SUBAPPLICATION Checkbox_TO_AD2_2 (* 2 VT-Checkboxes zu einer Bitmaske zusammenfassen und als AD2 (bidirektional) an einen Consumer weiterreichen (z.B. AOption_AD_DEMUX_2.K). Checkbox 1 -> Bit0, Checkbox 2 -> Bit1. Das vom Consumer zurueckgemeldete Echo (die tatsaechlich aktive Bitmaske) wird wieder auf die beiden Checkboxen zurueckgeschrieben. *)
  (* Standard: 61499-2; Description: Copyright (c) 2026 Meisterschulen am Ostbahnhof This program and the accompanying materials are made available under the terms of the Eclipse Public License 2.0 which is available at https://www.eclipse.org/legal/epl-2.0/ SPDX-License-Identifier: EPL-2.0 *)
  (* Version 1.0, 2026-10-13, Franz Höpfinger, Meisterschulen am Ostbahnhof, Ausgelagert aus Uebung_094b5_AX zur Wiederverwendung: Checkbox_IDA_TO_AX x2 + ASSEMBLE_AD_FROM_AX + AD_TO_AD2 + SPLIT_AD_INTO_AX + AX_TO_Checkbox x2. Fuer N=2 Bits/Checkboxes, analog zu AOption_AD_DEMUX_2. *)
  PACKAGE MyLib::sys;
  IMPORT isobus::UT::Q::const::IDs::ID_NULL;
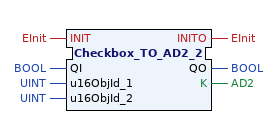
  EVENT_INPUT
    INIT : EInit; (* Initialization Request *)
  END_EVENT
  EVENT_OUTPUT
    INITO : EInit; (* Initialization Confirm *)
  END_EVENT
  VAR_INPUT
    QI : BOOL := TRUE; (* Quality Input - TRUE to enable service *)
    u16ObjId_1 : UINT := ID_NULL; (* Object ID Checkbox 1 (Bit0) *)
    u16ObjId_2 : UINT := ID_NULL; (* Object ID Checkbox 2 (Bit1) *)
  END_VAR
  VAR_OUTPUT
    QO : BOOL; (* Quality Output - TRUE if service executed successfully *)
  END_VAR
  PLUGS
    K : adapter::types::bidirectional::AD2;
  END_PLUGS
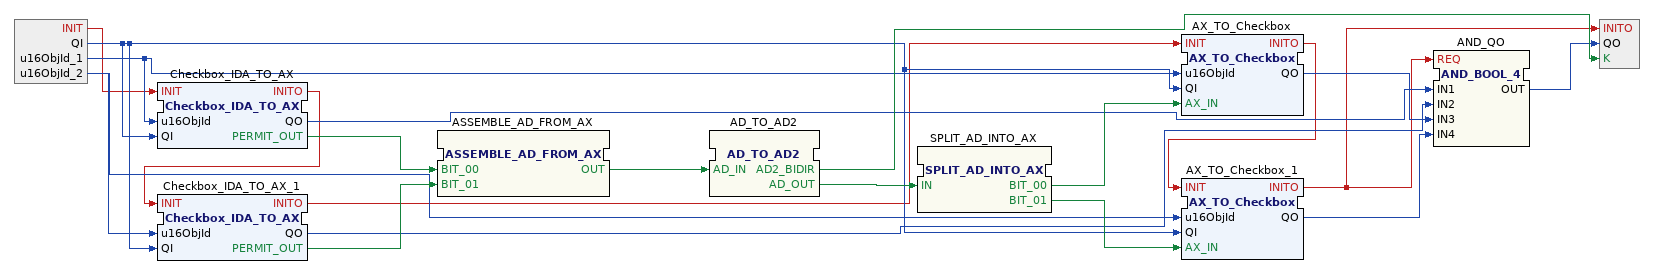
  FBS
    ASSEMBLE_AD_FROM_AX : adapter::assembling::ASSEMBLE_AD_FROM_AX;
    AD_TO_AD2 : adapter::conversion::bidirectional::AD_TO_AD2;
    SPLIT_AD_INTO_AX : adapter::splitting::SPLIT_AD_INTO_AX;
    AND_QO : iec61131::booleanOperators::AND_BOOL_4;
  END_FBS
  SUBAPPS
    Checkbox_IDA_TO_AX : MyLib::sys::Checkbox_IDA_TO_AX;
    Checkbox_IDA_TO_AX_1 : MyLib::sys::Checkbox_IDA_TO_AX;
    AX_TO_Checkbox : MyLib::sys::AX_TO_Checkbox;
    AX_TO_Checkbox_1 : MyLib::sys::AX_TO_Checkbox;
  END_SUBAPPS
  EVENT_CONNECTIONS
    INIT TO Checkbox_IDA_TO_AX.INIT;
    Checkbox_IDA_TO_AX.INITO TO Checkbox_IDA_TO_AX_1.INIT;
    Checkbox_IDA_TO_AX_1.INITO TO AX_TO_Checkbox.INIT;
    AX_TO_Checkbox.INITO TO AX_TO_Checkbox_1.INIT;
    AX_TO_Checkbox_1.INITO TO INITO;
    AX_TO_Checkbox_1.INITO TO AND_QO.REQ;
  END_CONNECTIONS
  DATA_CONNECTIONS
    u16ObjId_1 TO Checkbox_IDA_TO_AX.u16ObjId;
    u16ObjId_1 TO AX_TO_Checkbox.u16ObjId;
    u16ObjId_2 TO Checkbox_IDA_TO_AX_1.u16ObjId;
    u16ObjId_2 TO AX_TO_Checkbox_1.u16ObjId;
    QI TO Checkbox_IDA_TO_AX.QI;
    QI TO Checkbox_IDA_TO_AX_1.QI;
    QI TO AX_TO_Checkbox.QI;
    QI TO AX_TO_Checkbox_1.QI;
    Checkbox_IDA_TO_AX.QO TO AND_QO.IN1;
    Checkbox_IDA_TO_AX_1.QO TO AND_QO.IN2;
    AX_TO_Checkbox.QO TO AND_QO.IN3;
    AX_TO_Checkbox_1.QO TO AND_QO.IN4;
    AND_QO.OUT TO QO;
  END_CONNECTIONS
  ADAPTER_CONNECTIONS
    Checkbox_IDA_TO_AX.PERMIT_OUT TO ASSEMBLE_AD_FROM_AX.BIT_00;
    Checkbox_IDA_TO_AX_1.PERMIT_OUT TO ASSEMBLE_AD_FROM_AX.BIT_01;
    ASSEMBLE_AD_FROM_AX.OUT TO AD_TO_AD2.AD_IN;
    AD_TO_AD2.AD2_BIDIR TO K;
    AD_TO_AD2.AD_OUT TO SPLIT_AD_INTO_AX.IN;
    SPLIT_AD_INTO_AX.BIT_00 TO AX_TO_Checkbox.AX_IN;
    SPLIT_AD_INTO_AX.BIT_01 TO AX_TO_Checkbox_1.AX_IN;
  END_CONNECTIONS
END_SUBAPPLICATION
